(*
SPDX-FileCopyrightText: © 2026 Oleksandr Tiutyk <trofimich@gmail.com>
SPDX-License-Identifier: MIT
License: https://opensource.org/license/mit
*)

(*!
<summary>Reads a JSON document using scoped DOM handles.</summary>
<description>
Use a single instance from one task without reentry. UTF-8 text, including ASCII and empty strings, is decoded directly.
Legacy encodings use the native symbol converter.
</description>
*)

{attribute 'no_explicit_call' := 'do not call this function block directly'}
FUNCTION_BLOCK JsonConfigurationReader EXTENDS TOF_Core.Object IMPLEMENTS TOF_Core.IConfigurationReader
VAR_STAT
	_ClassName : STRING := __POUNAME();
END_VAR
VAR
	_Parser : Tc3_JsonXml.FB_JsonDomParser;
	_Converter : Tc3_JsonXml.FB_JsonReadWriteDatatype;
	_Value : TOF_Core.JSON_DOCUMENT;
END_VAR

(*!
<summary>Provides the concrete serializer class name.</summary>
<description>Borrows read-only instance storage that remains valid for the instance lifetime.</description>
*)
{attribute 'monitoring' := 'call'}
PROPERTY ClassName : REFERENCE TO STRING
GET
ClassName REF= _ClassName;
END_GET
END_PROPERTY

(*!
<summary>Attempts to find an optional object member without throwing.</summary>
<description>Returns EMPTY_NODE when absent. No exception escapes this method.</description>
<param name="node">Parent object node.</param>
<param name="name">Optional member field name.</param>
*)
METHOD FindField : TOF_Core.CONFIGURATION_NODE
VAR_INPUT
	node : TOF_Core.CONFIGURATION_NODE;
	name : STRING;
END_VAR
VAR
	member : __XWORD;
END_VAR
IF node.Handle = 0 OR_ELSE NOT _Parser.IsObject(v := node.Handle) THEN
	FindField := TOF_Core.ConfigurationNodes.EMPTY_NODE;
	RETURN;
END_IF

member := _Parser.FindMember(v := node.Handle, member := name);
FindField.Handle := member;
END_METHOD

(*!
<summary>Returns the number of elements of an array. Other shapes raise.</summary>
<description>
Use within one synchronous load. Handles borrow the active document and expire when it is replaced.
</description>
<param name="node">Array node.</param>
*)
METHOD GetArraySize : UDINT
VAR_INPUT
	node : TOF_Core.CONFIGURATION_NODE;
END_VAR
IF NOT IsArray(node := node) THEN
	throwInvalidDocumentException(reason := 'not an array', fieldName := '');
END_IF

GetArraySize := _Parser.GetArraySize(v := node.Handle);
END_METHOD

(*!
<summary>Finds a mandatory object member or raises.</summary>
<description>
Use within one synchronous load. Handles borrow the active document and expire when it is replaced.
</description>
<param name="node">Parent object node.</param>
<param name="name">Member field name.</param>
*)
METHOD GetField : TOF_Core.CONFIGURATION_NODE
VAR_INPUT
	node : TOF_Core.CONFIGURATION_NODE;
	name : STRING;
END_VAR
IF node.Handle = 0 OR_ELSE NOT _Parser.IsObject(v := node.Handle) THEN
	throwInvalidDocumentException(reason := 'not an object', fieldName := name);
END_IF

GetField.Handle := _Parser.FindMember(v := node.Handle, member := name);

IF GetField.Handle = 0 THEN
	throwInvalidDocumentException(reason := 'missing field', fieldName := name);
END_IF
END_METHOD

(*!
<summary>Returns an existing array item by zero-based index or raises.</summary>
<description>Use within one synchronous load. Out-of-bounds index raises an exception.</description>
<param name="node">Array node.</param>
<param name="index">Zero-based element index.</param>
*)
METHOD GetItem : TOF_Core.CONFIGURATION_NODE
VAR_INPUT
	node : TOF_Core.CONFIGURATION_NODE;
	index : UDINT;
END_VAR
IF NOT IsArray(node := node) THEN
	throwInvalidDocumentException(reason := 'not an array', fieldName := '');
END_IF

IF index >= _Parser.GetArraySize(v := node.Handle) THEN
	throwInvalidDocumentException(reason := 'index out of range', fieldName := '');
END_IF

GetItem.Handle := _Parser.GetArrayValueByIdx(v := node.Handle, idx := index);
END_METHOD

(*!
<summary>Reports whether the supplied value is an array.</summary>
<description>
Use within one synchronous load. Handles borrow the active document and expire when it is replaced.
</description>
<param name="node">Node to inspect.</param>
*)
METHOD IsArray : BOOL
VAR_INPUT
	node : TOF_Core.CONFIGURATION_NODE;
END_VAR
IsArray := node.Handle <> 0 AND_THEN _Parser.IsArray(v := node.Handle);
END_METHOD

(*!
<summary>Reports whether the supplied node refers to a present document element.</summary>
<description>Returns FALSE for an empty or unassigned node handle.</description>
<param name="node">Node to inspect.</param>
*)
METHOD IsPresent : BOOL
VAR_INPUT
	node : TOF_Core.CONFIGURATION_NODE;
END_VAR
IsPresent := node.Handle <> 0;
END_METHOD

(*!
<summary>Provides the compiler-initialized library namespace.</summary>
<description>Borrows read-only library storage; no allocation or ownership transfer occurs.</description>
*)
{attribute 'monitoring' := 'call'}
PROPERTY NamespaceName : REFERENCE TO STRING
GET
NamespaceName REF= CurrentNamespace.Name;
END_GET
END_PROPERTY

(*!
<summary>Parses a JSON configuration document and returns its root cursor node.</summary>
<description>Requires an object root. A new call invalidates all previously issued cursors.</description>
<param name="document">Null-terminated JSON document text.</param>
*)
METHOD Parse : TOF_Core.CONFIGURATION_NODE
VAR_IN_OUT CONSTANT
	document : TOF_Core.JSON_DOCUMENT;
END_VAR
Parse.Handle := _Parser.ParseDocument(sJson := document);

IF Parse.Handle = 0 THEN
	throwInvalidDocumentException(reason := 'parse failure', fieldName := '');
ELSIF NOT _Parser.IsObject(v := Parse.Handle) THEN
	throwInvalidDocumentException(reason := 'not an object', fieldName := '');
END_IF
END_METHOD

(*!
<summary>Reads one elementary value into a live typed destination or raises.</summary>
<description>
Use within one synchronous load. Handles borrow the active document and expire when it is replaced.
WSTRING requires a JSON string. Direct UTF-8 decoding checks the destination capacity before writing.
Native copy failures identify the operation and buffer size. Read the destination only after successful return.
</description>
<param name="node">Node containing the elementary value.</param>
<param name="valueType">Elementary IEC type class to decode.</param>
<param name="data">Writable pointer to the destination memory.</param>
<param name="size">Destination memory size in bytes.</param>
*)
METHOD ReadValue
VAR_INPUT
	node : TOF_Core.CONFIGURATION_NODE;
	valueType : TOF_Core.CONFIGURATION_VALUE_TYPE;
	data : PVOID;
	size : UDINT;
END_VAR
VAR
	typeName : STRING;
	target : POINTER TO STRING;
	result : HRESULT;
END_VAR
IF data = 0 OR_ELSE size = 0 THEN
	throwInvalidDocumentException(reason := 'type/size mismatch', fieldName := '');
END_IF

IF node.Handle = 0 THEN
	throwInvalidDocumentException(reason := 'missing field', fieldName := '');
END_IF

IF _Parser.IsNull(v := node.Handle)
	OR_ELSE _Parser.IsArray(v := node.Handle)
	OR_ELSE _Parser.IsObject(v := node.Handle)
THEN
	throwInvalidDocumentException(reason := 'type/size mismatch', fieldName := '');
END_IF

typeName := JsonDatatypes.ToDatatypeName(valueType := valueType, size := size);

IF typeName = '' THEN
	throwInvalidDocumentException(reason := 'type/size mismatch', fieldName := '');
END_IF

IF valueType = TOF_Core.CONFIGURATION_VALUE_TYPE.TYPE_STRING THEN
	target := data;

	IF NOT _Parser.IsString(v := node.Handle) THEN
		throwInvalidDocumentException(reason := 'type/size mismatch', fieldName := '');
	END_IF

	IF _Parser.CopyString(v := node.Handle, pStr := target^, nStr := size) = 0 THEN
		throwInvalidDocumentException(
			reason := TOF_Core.Strings.Concat255(
				'CopyString failed for ', typeName, ' (', TO_STRING(size), ' destination bytes)'
			),
			fieldName := ''
		);
	END_IF

	RETURN;
END_IF

IF valueType = TOF_Core.CONFIGURATION_VALUE_TYPE.TYPE_WSTRING THEN
	IF NOT _Parser.IsString(v := node.Handle) THEN
		throwInvalidDocumentException(reason := 'type/size mismatch', fieldName := '');
	END_IF

	IF readUtf8WideString(node := node, destination := data, size := size) THEN
		RETURN;
	END_IF
END_IF

IF _Parser.CopyJson(v := node.Handle, pDoc := _Value, nDoc := SIZEOF(_Value)) = 0 THEN
	throwInvalidDocumentException(
		reason := TOF_Core.Strings.Concat255(
			'CopyJson failed for ', typeName, ' (', TO_STRING(SIZEOF(_Value)), ' JSON buffer bytes)'
		),
		fieldName := ''
	);
END_IF

IF NOT _Converter.SetSymbolFromJson(
	sJson := _Value,
	sDatatype := typeName,
	nData := size,
	pData := data,
	hrErrorCode => result
) OR_ELSE result <> 0 THEN
	throwInvalidDocumentException(reason := 'parse failure', fieldName := '');
END_IF
END_METHOD

(*!
<summary>Reports the complete instance size in bytes.</summary>
<description>Uses XSIZEOF; separately allocated native resources are not included.</description>
*)
{attribute 'monitoring' := 'call'}
PROPERTY SelfSize : ULINT
GET
SelfSize := XSIZEOF(THIS^);
END_GET
END_PROPERTY

(*!
<summary>Decodes a JSON string directly into a WSTRING destination when its bytes are available as UTF-8.</summary>
<description>
Expects a live string node and a writable WSTRING buffer with a validated byte size. Returns FALSE
without writing when the copied text uses a legacy encoding.
The caller then uses the native symbol converter. Inspects JSON escapes before copying decoded text to an IEC string.
Both DOM and copy sizes include the terminator. Rejects a size mismatch,
an embedded null, insufficient destination capacity, or incomplete conversion. Conversion failure may modify the destination.
</description>
*)
METHOD PRIVATE readUtf8WideString : BOOL
VAR_INPUT
	node : TOF_Core.CONFIGURATION_NODE;
	destination : POINTER TO WSTRING;
	size : UDINT;
END_VAR
VAR
	// A JSON escape for U+0000, which IEC text cannot represent within a value.
	nullEscape : STRING(6) := '\u0000';
	jsonSize : UDINT;
	offset : UDINT;
	escapeIndex : UDINT;
	jsonBytes : POINTER TO BYTE;
	domStringSize : UDINT;
	copiedSize : UDINT;
	characterCount : UDINT;
	decodedCount : UDINT;
END_VAR
jsonSize := _Parser.CopyJson(v := node.Handle, pDoc := _Value, nDoc := SIZEOF(_Value));

IF jsonSize = 0 THEN
	throwInvalidDocumentException(reason := 'parse failure', fieldName := '');
END_IF

jsonBytes := ADR(_Value);
offset := 1; // Skip the opening JSON quote.

WHILE offset + SIZEOF(nullEscape) <= jsonSize DO
	IF jsonBytes[offset] = nullEscape[0] THEN
		escapeIndex := 1;

		WHILE escapeIndex < SIZEOF(nullEscape) - TOF_Core.Strings.CharSize
			AND_THEN jsonBytes[offset + escapeIndex] = nullEscape[escapeIndex]
		DO
			escapeIndex := escapeIndex + 1;
		END_WHILE

		IF escapeIndex = SIZEOF(nullEscape) - TOF_Core.Strings.CharSize THEN
			throwInvalidDocumentException(reason := 'parse failure', fieldName := '');
		END_IF

		// Skip the escaped byte as well, including a second backslash in a literal backslash pair.
		offset := offset + 1;
	END_IF

	offset := offset + 1;
END_WHILE

domStringSize := _Parser.GetStringLength(v := node.Handle);

copiedSize := _Parser.CopyString(v := node.Handle, pStr := _Value, nStr := SIZEOF(_Value));

IF copiedSize = 0
	OR_ELSE copiedSize <> domStringSize
	OR_ELSE TOF_Core.Strings.GetActualSize(value := _Value) <> copiedSize
THEN
	throwInvalidDocumentException(reason := 'parse failure', fieldName := '');
END_IF

IF copiedSize = TOF_Core.Strings.CharSize THEN
	destination^[0] := 0;
	readUtf8WideString := TRUE;
	RETURN;
END_IF

characterCount := Tc2_Utilities.UTF8Len(pUTF8 := ADR(_Value));

IF characterCount = 0 THEN
	RETURN;
END_IF

IF characterCount >= size / TOF_Core.WideStrings.CharSize THEN
	throwInvalidDocumentException(
		reason := TOF_Core.Strings.Concat255(
			'WSTRING needs ', TO_STRING(characterCount), ' characters, capacity ',
			TO_STRING(size / TOF_Core.WideStrings.CharSize - 1)
		),
		fieldName := ''
	);
END_IF

IF NOT Tc2_Utilities.UTF8_TO_WSTRING(
	pDstWSTRING := destination,
	pSrcUTF8 := ADR(_Value),
	nDstSize := size,
	nDstLen => decodedCount
) OR_ELSE decodedCount <> characterCount THEN
	throwInvalidDocumentException(reason := 'parse failure', fieldName := '');
END_IF

readUtf8WideString := TRUE;
END_METHOD

(*!
<summary>Reports an invalid or incompatible configuration value or document structure.</summary>
<description>
Constructs a diagnostic error message with the failure cause and optional member name, and raises StandardException.
The reader remains reusable by opening another document.
</description>
<param name="reason">Specific failure description.</param>
<param name="fieldName">Associated member field name, or empty when not applicable.</param>
*)
METHOD PRIVATE throwInvalidDocumentException
VAR_INPUT
	reason : STRING;
	fieldName : STRING;
END_VAR
VAR
	diagnosticMessage : TOF_Core.ERROR_MESSAGE;
END_VAR
IF fieldName <> '' THEN
	diagnosticMessage := TO_WSTRING(TOF_Core.Strings.Concat255(
		'Invalid JSON configuration: ',
		reason,
		' (field: ',
		fieldName,
		')'
	));
ELSE
	diagnosticMessage := TO_WSTRING(TOF_Core.Strings.Concat255('Invalid JSON configuration: ', reason));
END_IF

TOF_Core.Exceptions.ThrowStandard(
	sourceNamespaceName := NamespaceName,
	sourceClassName := ClassName,
	sourcePOUName := __POUNAME(),
	sourcePosition := __POSITION(),
	message := diagnosticMessage,
	errorCode := 16#80070057
);
END_METHOD

END_FUNCTION_BLOCK

(* stored: Version 1.1.0.1
   POU JsonConfigurationReader: Id {236a8e5c-23da-49c0-8af5-0fa696e16ceb}, SpecialFunc None
   Folder Service methods: Id {bec439dc-2b8a-4719-bfbc-2186f8994348}
   Property ClassName: Id {cb3e6f75-e064-4b44-9538-0a7bd332335c}
   Get Get: Id {512664b3-26d4-4b25-8af0-39c7b7d2485a}
   Method FindField: Id {cd757efd-cff4-4b37-b363-1b9042c90708}
   Method GetArraySize: Id {49417c52-e7f4-414e-92d2-72a8f1d07e48}
   Method GetField: Id {b6f25c33-3a9f-4d17-b447-fe531a426ea2}
   Method GetItem: Id {6d689d67-8cfe-4aac-b45f-4635cb27afba}
   Method IsArray: Id {91240330-ce82-4217-ad18-08ada72cf717}
   Method IsPresent: Id {6af041a0-5276-4f46-9640-1ea64cfd1a53}
   Property NamespaceName: Id {ed4f9045-a704-45f7-9e75-4d04cfcac736}
   Get Get: Id {f1a7faa9-09f0-4b68-81b8-f301754cf572}
   Method Parse: Id {458f1032-13e5-4c9a-9aa5-8b26b6414885}
   Method ReadValue: Id {ce16e1f6-9681-4b51-a5a6-ee3bdb56e190}
   Property SelfSize: Id {e1ba1bb4-ae22-42ad-8dba-e61c26974727}
   Get Get: Id {38e6e3a8-2e64-402d-9fcd-d603b0515426}
   Method readUtf8WideString: Id {80593a06-c9e1-4f7e-9300-d6f64d094430}
   Method throwInvalidDocumentException: Id {e0005382-6117-4a05-a35e-b58f52a8f44d} *)
